Fanuc KAREL source: ko00096.KL

-- PROVISIONAL review KL for V1013-1; original PC SHA256 7e1b6d768918382d26f41a114b921a05b7497cfb19768d750f75d7ddeab8b50e
-- Incomplete behavior may be omitted. Consult companion uncertainty JSON. Do not deploy.
PROGRAM KO00096
%NOLOCKGROUP
BEGIN
  -- UNRESOLVED_PC offsets 5-12; opcodes 9D,23
  -- UNRESOLVED_PC offsets 17-69; opcodes 27,27,49,7E,AD,27,49,7E,AD,22,31,7E,4A
  -- UNRESOLVED_PC offsets 74-78; opcodes 7F
END KO00096
